Fanuc KAREL source: kb00010.KL

-- PROVISIONAL review KL for V940-1; original PC SHA256 df257b8981e6df1bf385aa0dff56a5560db194c4603773315e14451a8c4ed0e2
-- Incomplete behavior may be omitted. Consult companion uncertainty JSON. Do not deploy.
PROGRAM KB00010
%NOLOCKGROUP
BEGIN
  -- V9_ZERO_TABLE_METADATA_HINT layout=0002_ascii; no indexed target words; source/name/runtime held
  -- UNRESOLVED_PC offsets 5-14; opcodes 3F,75
  -- UNRESOLVED_PC offsets 19-28; opcodes 3F,75
  -- UNRESOLVED_PC offsets 33-40; opcodes 9D,23
  -- UNRESOLVED_PC offsets 45-52; opcodes 9D,23
  -- UNRESOLVED_PC offsets 57-66; opcodes 3F,75
  -- UNRESOLVED_PC offsets 71-78; opcodes 9D,23
  -- UNRESOLVED_PC offsets 83-129; opcodes 27,22,2A,22,2A,22,22,22,2A,22,31
  -- UNRESOLVED_PC offsets 134-138; opcodes 7F
END KB00010
